//{attribute 'qualified_only'}
VAR_GLOBAL
	stVisuPLC_To_PLC		AT %MB1000 : ST_VisuPLC_To_PLC;
	stPLC_To_VisuPLC		AT %MB2000 : ST_PLC_To_VisuPLC;
	
	i_stVisuPLC_To_PLC		AT %I* : ST_VisuPLC_To_PLC;
	q_stPLC_To_VisuPLC		AT %Q* : ST_PLC_To_VisuPLC;	
END_VAR

(* stored: Version 1.1.0.1, ProductVersion 3.1.4024.15
   GVL g_HMI_Panel: Id {f85eecbd-41e4-462b-af15-59cdbfb1c9a3} *)
